// TIA Portal V17 export
// export: Created 2026-11-08T05:50:29.4104014Z, ExportSetting WithDefaults, DisplayName Totally Integrated Automation Portal, DisplayVersion V17, DisplayName TIA Portal Openness, DisplayVersion V17, DisplayName TIA Portal Version Control Interface, DisplayVersion V17, DisplayName STEP 7 Professional, DisplayVersion V17, DisplayName STEP 7 Safety, DisplayVersion V17, DisplayName WinCC Professional, DisplayVersion V17
VAR_GLOBAL   // PLC tag table "Motores"
   KM1_Motor AT %M10.3 : Bool;   // Contactor KM1 del motor M1
   MOT1_Termico_Falla AT %M10.2 : Bool;   // Relé térmico M1: 1 = disparado
END_VAR
